Staubli VAL3: HMI_prog.pjx

--- HMI_prog.pjx ---
Parameters version=s8.15.1Cs9_BS3177 stackSize=5000 millimeterUnit=true
Program file=bind.pgx
Program file=bind_edit.pgx
Program file=main.pgx
Program file=onSimulate.pgx
Program file=onStart.pgx
Program file=refreshlist.pgx
Program file=refreshproglist.pgx
Program file=selEndProg.pgx
Program file=selMainProg.pgx
Program file=selStartUpProg.pgx
Program file=start.pgx
Program file=stop.pgx
Data file=HMI_prog.dtx
Library alias=program path=Disk://source/projectSource/program/program.pjx
Library alias=util path=Disk://HMI_cs9/HMI_util/HMI_util.pjx
Library alias=trajectory path=Disk://source/projectSource/trajectory/trajectory.pjx
Library alias=actionData path=Disk://data/actionData/actionData.pjx
Library alias=simulate path=Disk://HMI_cs9/simulate/simulate.pjx
Library alias=editprog path=Disk://HMI_cs9/HMI_progEdit/HMI_progEdit.pjx
Library alias=progTemp path=Disk://source/template/progTemp/progTemp.pjx
Library alias=rs path=Disk://source/projectSource/robotStatus/robotStatus.pjx

--- HMI_prog.dtx ---
string sProgLsit
num nPageIndex
num nPageNum
string sSelProg
string sPageIndex
string sPageNum
public bool bBool[10]
bool bToSave
bool bBack
public bool bEditBool[9]
string sEditIndex
string sEditPage
string sSelTRAJ
num nEditPage
num nEditIndex
string sList[49]
bool bEditBack
bool bInsert
bool bCancel
string sSelType
string sSelItem
string sLastType
string sInsertList
num nType
public string sIF_Type[3]
public string sIF_Index[3]
num nIF_value[3]
num nProgType
string sInitialPassword = "55582930"

--- main.pgx ---
public program main()
  local bool l_bExit
  local bool l_bRefresh
  local bool l_bResult
  local string l_sEntryPassword
begin
  do
    if util:sPage!="prog"
      util:sPage="prog"
      call onStart()
      call bind()
      userPage(util:sPage)
      delay(0.5)
      l_bRefresh=true
    endIf

    if bBool[0]
      bBool[0]=false
      //新建
      call program:new(bToSave)
      l_bRefresh=true
    elseIf bBool[1]
      bBool[1]=false
      //编辑
      if bToSave
        bToSave=false
        call program:onSave(bToSave)
      endIf
      if sSelProg!=""
        call editprog:main(sSelProg)
      else
        userPageAlert("未选择有效项")
      endIf
      l_bRefresh=true
    elseIf bBool[2]
      bBool[2]=false
      //删除
      if find(sSelProg,"prod")!=-1
        //ADD BY Liuzhengang20260225
        l_bResult=userPagePrompt("请输入密码",l_sEntryPassword)
        if l_bResult==false
          return
        else
          if l_sEntryPassword!=sInitialPassword[0]
            popUpMsg("密码错误")
            return
          else
            call program:deleteProg(sSelProg,bToSave)
            l_bRefresh=true
          endIf
        endIf
        //        userPageAlert("不可删除选项！")
        //        return
      else
        call program:deleteProg(sSelProg,bToSave)
        l_bRefresh=true
      endIf

    elseIf bBool[3]
      bBool[3]=false
      //保存
      call program:onSave(bToSave)
    elseIf bBool[4]
      bBool[4]=false
      //复制
      l_bRefresh=true
      call program:copy(sSelProg,bToSave)
    elseIf bBool[5]
      bBool[5]=false
      call simulate:simulatePROG(sSelProg)
    elseIf bBool[6]
      bBool[6]=false
      nPageIndex=0
      l_bRefresh=true
    elseIf bBool[7]
      bBool[7]=false
      if nPageIndex>0
        nPageIndex=nPageIndex-1
        l_bRefresh=true
      endIf

    elseIf bBool[8]
      bBool[8]=false
      if nPageIndex<nPageNum-1
        nPageIndex=nPageIndex+1
        l_bRefresh=true
      endIf
    elseIf bBool[9]
      bBool[9]=false
      nPageIndex=nPageNum-1
      l_bRefresh=true
    elseIf bBack
      bBack=false
      if bToSave
        bToSave=false
        l_bResult=userPageConfirm("是否保存数据")
        if l_bResult
          call program:onSave(bToSave)
        endIf
      endIf
      l_bExit=true
    endIf

    if l_bRefresh
      l_bRefresh=false
      // call program:getProgList(sProgLsit)
      call refreshlist()
      // userPageBind("prog","lst1","options",sProgLsit,size(sProgLsit),"r")
      // call refreshproglist()
    endIf


    delay(0)
  until l_bExit==true
end

--- start.pgx ---
program start()
begin
end

--- bind.pgx ---
public program bind()
  local num l_i
  local string l_sbtn
begin
  //lst
  userPageBind("prog","lst1","options",sList,49,"r")
  userPageBind("prog","lst1","value",sSelProg,1,"rw")
  for l_i = 0 to size(bBool)-1
    l_sbtn="btn"+toString("",l_i)
    userPageBindClick("prog",l_sbtn,bBool[l_i],true)
  endFor
  userPageBindClick("prog","btnback",bBack,true)
  userPageBind("prog","lbleditindex","innerHTML",sPageIndex,1,"r")
  userPageBind("prog","lbleditpage","innerHTML",sPageNum,1,"r")
end

--- bind_edit.pgx ---
program bind_edit()
  local num l_i
  local string l_sbtn
begin
  for l_i = 0 to size(bEditBool)-1
    l_sbtn="btn"+toString("",l_i)
    userPageBindClick("editProg",l_sbtn,bEditBool[l_i],true)
  endFor

  userPageBindClick("editProg","btnback",bEditBack,true)

  userPageBind("editProg","lbleditindex","innerHTML",sEditIndex,1,"r")
  userPageBind("editProg","lbleditpage","innerHTML",sEditPage,1,"r")

  userPageBind("editProg","lst1","value",sSelTRAJ,1,"rw")
end

--- onSimulate.pgx ---
public program onSimulate()
begin
end

--- onStart.pgx ---
public program onStart()
  local num l_nResult
begin
  // call program:loadPROG(0,l_nResult)
  //  if l_nResult!=0
  //    popUpMsg("库加载错误："+toString("",l_nResult))
  //  endIf

  // call refreshproglist()
  call program:getProgList(sProgLsit)
  call refreshlist()

  nPageIndex=0
  nPageNum=roundUp(size(sProgLsit)/49)

  if !isDefined(progTemp:pProgItem[sSelProg])
    sSelProg=""
  endIf
  //
  sPageIndex=toString("",nPageIndex+1)
  sPageNum=toString("",nPageNum)
end

--- refreshlist.pgx ---
public program refreshlist()
  local string l_skey
  local num l_i
  local num l_nSize
begin
  call program:getProgList(sProgLsit)
  l_nSize=size(sProgLsit)

  if l_nSize<=49
    nPageNum=1
  else
    nPageNum=roundUp(l_nSize/49)
  endIf

  if nPageNum==1
    for l_i = 0 to size(sList)-1
      sList[l_i]=""
    endFor
    for l_i = 0 to l_nSize-1
      sList[l_i]=sProgLsit[l_i]
    endFor
  else
    if nPageIndex<nPageNum-1
      for l_i = 0 to 48
        sList[l_i]=sProgLsit[49*nPageIndex+l_i]
      endFor
    else
      for l_i = 0 to size(sList)-1
        sList[l_i]=""
      endFor
      for l_i = 0 to(l_nSize%49)-1
        sList[l_i]=sProgLsit[49*nPageIndex+l_i]
      endFor
    endIf
  endIf
  userPageBind("prog","lst1","options",sList,size(sList),"r")
  sPageIndex=toString("",nPageIndex+1)
  sPageNum=toString("",nPageNum)
end

--- refreshproglist.pgx ---
public program refreshproglist()
  local num l_nSize
  local num l_nProgSize
  local num l_i
  local string l_sMsg
begin
  call program:getProgItemSize(sSelProg,l_nProgSize)
  if l_nProgSize<50
    nEditPage=1
  else
    nEditPage=roundUp(l_nProgSize/49)
  endIf

  if nEditIndex>(nEditPage-1)
    nEditIndex=(nEditPage-1)
  endIf
  //slist
  if nEditIndex==(nEditPage-1)
    if l_nProgSize%49==0
      l_nSize=49
    else
      l_nSize=l_nProgSize%49
    endIf
    for l_i = 0 to l_nSize-1
      call program:pointToString(l_sMsg,sSelProg,l_i+49*nEditIndex)
      sList[l_i]=toString("",l_i+49*nEditIndex)+l_sMsg
    endFor
    if l_nSize<49
      for l_i= l_nSize to size(sList)-1
        sList[l_i]=""
      endFor
    endIf
  else
    for l_i = 0 to size(sList)-1
      call program:pointToString(l_sMsg,sSelProg,l_i+49*nEditIndex)
      sList[l_i]=toString("",l_i+49*nEditIndex)+l_sMsg
    endFor
  endIf
  userPageBind("prog","lst1","options",sList,size(sList),"r")
  sEditIndex=toString("",nEditIndex+1)
  sEditPage=toString("",nEditPage)

end

--- selEndProg.pgx ---
public program selEndProg()
begin
  nProgType=1
end

--- selMainProg.pgx ---
public program selMainProg()
begin
  nProgType=2
end

--- selStartUpProg.pgx ---
public program selStartUpProg()
begin
  nProgType=1
end

--- stop.pgx ---
program stop()
begin
end
